(* IEC 61131-3 sources: rusty/tests/lit/cfc/blocks/method_call, 2 files *)

(* ---- main.st ---- *)
FUNCTION main : DINT
    method_call();
    method_call();
    // CHECK: result = 6, doubled = 12
    printf('result = %d, doubled = %d$N', method_call.result, method_call.dbl);
END_FUNCTION

(* ---- counter.st ---- *)
FUNCTION_BLOCK counter
VAR
    count : DINT;
END_VAR
METHOD bump : DINT
VAR_INPUT
    step : DINT;
END_VAR
VAR_OUTPUT
    doubled : DINT;
END_VAR
    count := count + step;
    doubled := count * 2;
    bump := count;
END_METHOD
END_FUNCTION_BLOCK
